Fanuc KAREL source: kt00745.KL

-- PROVISIONAL review KL for V940-1; original PC SHA256 92b77fe70471aa01d1e440d6f6259a25764e796ebc43607f4f62bd73bd558775
-- Incomplete behavior may be omitted. Consult companion uncertainty JSON. Do not deploy.
PROGRAM KT00745
%NOLOCKGROUP
BEGIN
  -- V9_ZERO_TABLE_METADATA_HINT layout=0001; no indexed target words; source/name/runtime held
  -- UNRESOLVED_PC offsets 5-18; opcodes 22,1D,23
  -- UNRESOLVED_PC offsets 23-27; opcodes 7F
END KT00745
